Fanuc KAREL source: KA00064.KL

PROGRAM KA00064
%NOLOCKGROUP
VAR
  SRC: XYZWPR
  DST: STRING[80]
BEGIN
  SRC.X = 1.0
  DST = SRC
END KA00064
